Fanuc KAREL source: KO00012.KL

PROGRAM KO00012
%NOLOCKGROUP
VAR
  P1: XYZWPR
  P2: XYZWPR
  P3: XYZWPR
  OUT: JOINTPOS
BEGIN
  OUT = FRAME(P1, P2, P3)
END KO00012
